(* IEC 61131-3 sources: trust-platform/manual-tests/clean/src, 1 file *)

(* ---- DebugMain.st ---- *)
PROGRAM DebugMain
VAR
    x : DINT := 1;
    y : DINT := 2;
    sum : DINT;
END_VAR

sum := x + y;
END_PROGRAM
